FUNCTION_BLOCK NextFeedHorizonDiag (* CAT Function Block Type *)
  (* Standard: 61499-2 *)
  (* Version 0.0, 10/6/2026, Schneider Electric, template *)
  PACKAGE SE.Nereda;
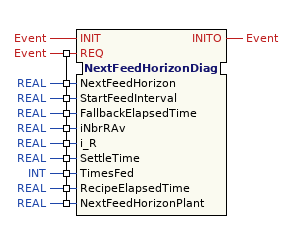
  EVENT_INPUT
    INIT; (* Initialization Request *)
    REQ WITH NextFeedHorizon, StartFeedInterval, FallbackElapsedTime, i_R, SettleTime, iNbrRAv, TimesFed, RecipeElapsedTime, NextFeedHorizonPlant; (* Normal Execution Request *)
  END_EVENT
  EVENT_OUTPUT
    INITO; (* Initialization Confirm *)
  END_EVENT
  VAR_INPUT
    NextFeedHorizon : REAL;
    StartFeedInterval : REAL;
    FallbackElapsedTime : REAL;
    iNbrRAv : REAL;
    i_R : REAL;
    SettleTime : REAL;
    TimesFed : INT;
    RecipeElapsedTime : REAL;
    NextFeedHorizonPlant : REAL;
  END_VAR
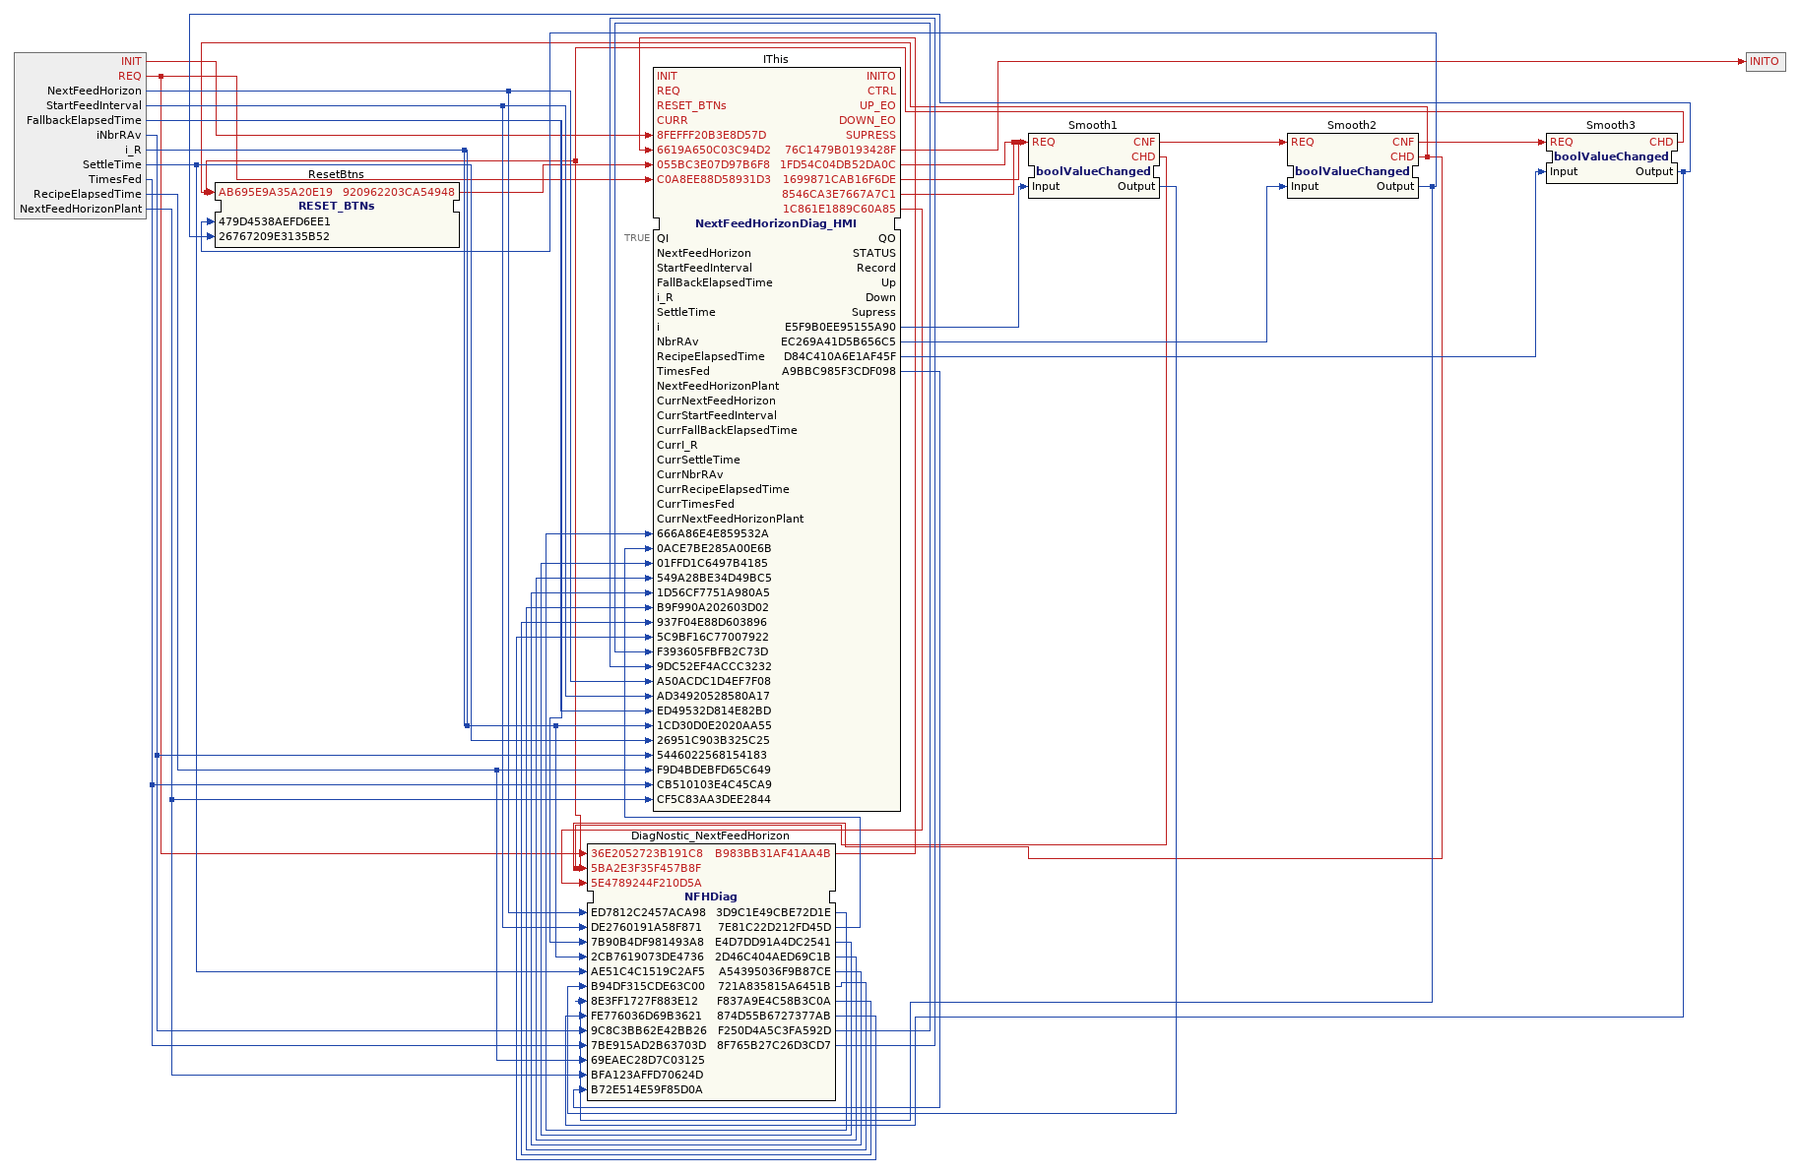
  FBS
    DiagNostic_NextFeedHorizon : NFHDiag;
    IThis : NextFeedHorizonDiag_HMI(QI := TRUE);
    ResetBtns : RESET_BTNs;
    Smooth1 : boolValueChanged;
    Smooth2 : boolValueChanged;
    Smooth3 : boolValueChanged;
  END_FBS
  EVENT_CONNECTIONS
    REQ TO DiagNostic_NextFeedHorizon.36E2052723B191C8;
    Smooth1.CNF TO Smooth2.REQ;
    Smooth2.CNF TO Smooth3.REQ;
    Smooth1.CHD TO DiagNostic_NextFeedHorizon.5BA2E3F35F457B8F;
    Smooth2.CHD TO DiagNostic_NextFeedHorizon.5BA2E3F35F457B8F;
    Smooth3.CHD TO DiagNostic_NextFeedHorizon.5BA2E3F35F457B8F;
    Smooth2.CHD TO ResetBtns.AB695E9A35A20E19;
    Smooth3.CHD TO ResetBtns.AB695E9A35A20E19;
    INIT TO IThis.8FEFFF20B3E8D57D;
    DiagNostic_NextFeedHorizon.B983BB31AF41AA4B TO IThis.6619A650C03C94D2;
    ResetBtns.920962203CA54948 TO IThis.055BC3E07D97B6F8;
    REQ TO IThis.C0A8EE88D58931D3;
    IThis.76C1479B0193428F TO INITO;
    IThis.1FD54C04DB52DA0C TO Smooth1.REQ;
    IThis.1699871CAB16F6DE TO Smooth1.REQ;
    IThis.8546CA3E7667A7C1 TO Smooth1.REQ;
    IThis.1C861E1889C60A85 TO DiagNostic_NextFeedHorizon.5E4789244F210D5A;
  END_CONNECTIONS
  DATA_CONNECTIONS
    NextFeedHorizon TO DiagNostic_NextFeedHorizon.ED7812C2457ACA98;
    StartFeedInterval TO DiagNostic_NextFeedHorizon.DE2760191A58F871;
    FallbackElapsedTime TO DiagNostic_NextFeedHorizon.7B90B4DF981493A8;
    i_R TO DiagNostic_NextFeedHorizon.2CB7619073DE4736;
    SettleTime TO DiagNostic_NextFeedHorizon.AE51C4C1519C2AF5;
    Smooth1.Output TO DiagNostic_NextFeedHorizon.B94DF315CDE63C00;
    Smooth2.Output TO DiagNostic_NextFeedHorizon.8E3FF1727F883E12;
    Smooth2.Output TO ResetBtns.479D4538AEFD6EE1;
    Smooth3.Output TO DiagNostic_NextFeedHorizon.FE776036D69B3621;
    Smooth3.Output TO ResetBtns.26767209E3135B52;
    iNbrRAv TO DiagNostic_NextFeedHorizon.9C8C3BB62E42BB26;
    TimesFed TO DiagNostic_NextFeedHorizon.7BE915AD2B63703D;
    RecipeElapsedTime TO DiagNostic_NextFeedHorizon.69EAEC28D7C03125;
    NextFeedHorizonPlant TO DiagNostic_NextFeedHorizon.BFA123AFFD70624D;
    DiagNostic_NextFeedHorizon.3D9C1E49CBE72D1E TO IThis.666A86E4E859532A;
    DiagNostic_NextFeedHorizon.7E81C22D212FD45D TO IThis.0ACE7BE285A00E6B;
    DiagNostic_NextFeedHorizon.E4D7DD91A4DC2541 TO IThis.01FFD1C6497B4185;
    DiagNostic_NextFeedHorizon.2D46C404AED69C1B TO IThis.549A28BE34D49BC5;
    DiagNostic_NextFeedHorizon.A54395036F9B87CE TO IThis.1D56CF7751A980A5;
    DiagNostic_NextFeedHorizon.721A835815A6451B TO IThis.B9F990A202603D02;
    DiagNostic_NextFeedHorizon.F837A9E4C58B3C0A TO IThis.937F04E88D603896;
    DiagNostic_NextFeedHorizon.874D55B6727377AB TO IThis.5C9BF16C77007922;
    DiagNostic_NextFeedHorizon.F250D4A5C3FA592D TO IThis.F393605FBFB2C73D;
    DiagNostic_NextFeedHorizon.8F765B27C26D3CD7 TO IThis.9DC52EF4ACCC3232;
    NextFeedHorizon TO IThis.A50ACDC1D4EF7F08;
    StartFeedInterval TO IThis.AD34920528580A17;
    FallbackElapsedTime TO IThis.ED49532D814E82BD;
    i_R TO IThis.1CD30D0E2020AA55;
    SettleTime TO IThis.26951C903B325C25;
    iNbrRAv TO IThis.5446022568154183;
    RecipeElapsedTime TO IThis.F9D4BDEBFD65C649;
    TimesFed TO IThis.CB510103E4C45CA9;
    NextFeedHorizonPlant TO IThis.CF5C83AA3DEE2844;
    IThis.E5F9B0EE95155A90 TO Smooth1.Input;
    IThis.EC269A41D5B656C5 TO Smooth2.Input;
    IThis.D84C410A6E1AF45F TO Smooth3.Input;
    IThis.A9BBC985F3CDF098 TO DiagNostic_NextFeedHorizon.B72E514E59F85D0A;
  END_CONNECTIONS
END_FUNCTION_BLOCK
